Fanuc KAREL source: kt00585.KL

-- PROVISIONAL review KL for V770-1; original PC SHA256 5b7fd4b3f0cacac7b25b167750c26e3d1ed21c79ea2527283a43ab1ab064fa80
-- Incomplete behavior may be omitted. Consult companion uncertainty JSON. Do not deploy.
PROGRAM KT00585
%NOLOCKGROUP
VAR
  I1 : INTEGER
-- UNRESOLVED_DECL V2 type=000013
-- UNRESOLVED_DECL OUT type=000013
BEGIN
  -- UNRESOLVED_PC offsets 5-16; opcodes 2E,23
  -- UNRESOLVED_PC offsets 21-36; opcodes 2E,22,32,35
  -- UNRESOLVED_PC offsets 41-63; opcodes 21,49,8B,4A
  -- UNRESOLVED_PC offsets 68-72; opcodes 7F
END KT00585
